TYPE ST_PolarIIChamber_OpenCloseServiceStatus :
STRUCT
	Open : ST_ServiceStatus;
	Close : ST_ServiceStatus;
END_STRUCT
END_TYPE

(* stored: Version 1.1.0.1, ProductVersion 3.1.4026.18
   DUT ST_PolarIIChamber_OpenCloseServiceStatus: Id {14000000-0000-0000-0000-000000000036} *)
